(* PLC project probe.project, CODESYS CODESYS V3.5 SP17 Patch 3 *)
(* stored: creationDateTime 2026-10-20T03:54:26.7557386, modificationDateTime 1601-01-01T03:00:00 *)

FUNCTION_BLOCK FB_ProbeFbd
  VAR_INPUT
    rLevel : REAL;
    rHigh : REAL;
    xEnable : BOOL;
    xAck : BOOL;
  END_VAR
  VAR_OUTPUT
    xOut : BOOL;
  END_VAR
  VAR
    xHigh : BOOL;
    xAlarm : BOOL;
  END_VAR

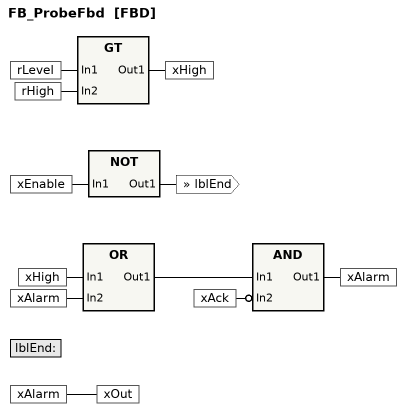
(* FBD diagram, written out as Structured Text *)
xHigh := rLevel > rHigh;
(* --- network: Пропуск при отключении --- *)
IF NOT xEnable THEN JMP lblEnd; END_IF;
(* --- network: Защёлка тревоги --- *)
xAlarm := (xHigh OR xAlarm) AND NOT xAck;
lblEnd:
(* --- network: Выход --- *)
xOut := xAlarm;
END_FUNCTION_BLOCK
